TYPE "ST_PressDemoStationCfg"
VERSION : 0.1
   STRUCT
      SchemaVersion : UInt := 2;
      DegradationPercent : UInt := 10;
      RequireTwoHandStart : Bool := TRUE;
   END_STRUCT;

END_TYPE

